// TIA Portal V21 export
// export: Created 2026-11-11T00:47:52.0382398Z, ExportSetting WithDefaults, DisplayName Totally Integrated Automation Portal, DisplayVersion V21 Update 3, DisplayName STEP 7 Professional, DisplayVersion V21 Update 3, DisplayName STEP 7 Safety, DisplayVersion V21, DisplayName Tech WebApplication, DisplayVersion V21, DisplayName WinCC Basic/Comfort/Advanced, DisplayVersion V21 Update 3, DisplayName WinCC Unified, DisplayVersion V21 Update 3
FUNCTION_BLOCK "FB_Lad_Trcv"   // FB350, LAD
{ S7_Optimized_Access := 'TRUE' }
VERSION : 0.1
// stored: AutoNumber true, IsIECCheckEnabled false, IsRetainMemResEnabled false, MemoryReserve 100, SetENOAutomatically false, UDAEnableTagReadback false
   VAR_INPUT
      en_r : Bool;
      cont : Bool;
      len : UInt;
      id : CONN_OUC;
      adhoc : Bool;
   END_VAR
   VAR_OUTPUT
      done : Bool;
      busy : Bool;
      err : Bool;
      status : Word;
      rcvdlen : UInt;
   END_VAR
   VAR_IN_OUT
      connect : TCON_IP_v4;
      data : Array[0..99] of Byte;
      comrst : Bool;
      addr : Variant;
   END_VAR
   VAR
      inst { S7_SetPoint := 'True'} : TRCV;
   END_VAR
BEGIN

REGION Network 1: TRCV
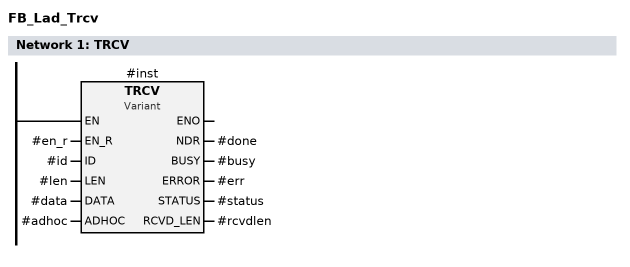
   RUNG wire#powerrail
      { S7_Templates := "[card := 1, ptr_type := Variant, value_type := UDInt, id_type := CONN_OUC]" } #inst.TRCV(EN_R := #en_r, ID := #id, LEN := #len, NDR => #done, BUSY => #busy, ERROR => #err, STATUS => #status, RCVD_LEN => #rcvdlen, DATA := #data, ADHOC := #adhoc)
   END_RUNG
   // the same network as SCL:
   #inst(EN_R := #en_r,   // TRCV
         ID := #id,
         LEN := #len,
         DATA := #data,
         ADHOC := #adhoc,
         NDR => #done,
         BUSY => #busy,
         ERROR => #err,
         STATUS => #status,
         RCVD_LEN => #rcvdlen);
END_REGION
END_FUNCTION_BLOCK
